  rq_init_comm_if_connected(9, "1")
  rq_init_comm_if_connected(2, "2")
  rq_init_comm_if_connected(3, "3")
  rq_init_comm_if_connected(4, "4")
  rq_print_connected_grippers()
  rq_gripper_communication_thread = run rq_gripper_communication()
  set_closed_norm(97.6470588235294, "1")
  set_open_norm(1.1764705882352942, "1")
  set_closed_mm(0.0, "1")
  set_open_mm(53.0, "1")
  set_closed_norm(100.0, "2")
  set_open_norm(0.0, "2")
  set_closed_mm(0.0, "2")
  set_open_mm(50.0, "2")
  set_closed_norm(100.0, "3")
  set_open_norm(0.0, "3")
  set_closed_mm(0.0, "3")
  set_open_mm(50.0, "3")
  set_closed_norm(100.0, "4")
  set_open_norm(0.0, "4")
  set_closed_mm(0.0, "4")
  set_open_mm(50.0, "4")
  rq_current_limit_enabled = False
  while(not rq_gripper_communication_thread_started):
      sleep(0.008)
  end
  # end: URCap Installation Node
  step_count_126a9c52_0873_4ea5_a9d9_3503bc14fb30 = 0.0
  thread Step_Counter_Thread_0450802b_b3f4_44ca_aa13_af17d282832f():
    while (True):
      step_count_126a9c52_0873_4ea5_a9d9_3503bc14fb30 = step_count_126a9c52_0873_4ea5_a9d9_3503bc14fb30 + 1.0
      sync()
    end
  end
  run Step_Counter_Thread_0450802b_b3f4_44ca_aa13_af17d282832f()
  global TMR_Barcode=0
  global TMR_Barcode_is_counting=False
  thread Timer_Thread():
    while (True):
      if (TMR_Barcode_is_counting):
        TMR_Barcode = TMR_Barcode + get_steptime()
      end
      sync()
    end
  end
  run Timer_Thread()
  $ 2 "BeforeStart"
  $ 3 "Before start"
  $ 4 "Script: SCRIPT Transitions V6.6.script"
  #*****************************************************
  # customer          :   INTERNAL
  # project name      :
  #****************************************************
  # controller        :   UR
  # software          :   5.13
  #****************************************************
  # author            :   P. Koehnke
  # Copyright (c)     :   United Robotics Group
  #                       An der Riede 2
  #                       28816 Stuhr
  #                       Germany
  #****************************************************
  # description       :   transition between workareas
  # version:      	:   1.2
  # created           :   28.02.2024
  # updated           :
  #****************************************************
  # modifications     :
  #
  # date              :
  # name              :
  # reason            :
  #****************************************************

  ######################### further development #########################
  #   - that the robot can switch the configuration, if necessary
  #   - introduction of structs
  #######################################################################

  ######################### to be adjusted #########################
  local WORKAREA_1 = [-0.280,-0.680,-0.001, 0.280, 0.100, 1.000]    # workarea 1 (platform)
  local WORKAREA_2 = [-1.000,-1.000,-1.000,-0.290, 0.100, 1.000]    # workarea 2 (front right)
  local WORKAREA_3 = [-1.000, 0.100,-1.000, 0.000, 1.000, 1.000]    # workarea 3 (back right)
  local WORKAREA_4 = [ 0.000, 0.100,-1.000, 1.000, 1.000, 1.000]    # workarea 4 (back left)
  local WORKAREA_5 = [ 0.290,-1.000,-1.000, 1.000, 0.100, 1.000]    # workarea 5 (front left)
  local WORKAREA_6 = [-0.290,-1.000,-1.000, 0.290,-0.560, 1.000]    # workarea 6 (front front)
  local WORKAREA_7 = [0,0,0,0,0,0]    # reserved
  local WORKAREA_8 = [0,0,0,0,0,0]    # reserved
  local WORKAREA_9 = [0,0,0,0,0,0]    # reserved
  local WORKAREA_10 = [0,0,0,0,0,0]   # reserved

  local PSE_WA_1 = p[ 0.000,-0.450, 0.300, 0.000, 0.000, 0.000]
  local PSE_WA_2 = p[-0.300,-0.300, 0.300, 0.000, 0.000, d2r(-90)]
  local PSE_WA_3 = p[-0.300, 0.300, 0.300, 0.000, 0.000, d2r(-135)]
  local PSE_WA_4 = p[ 0.300, 0.300, 0.300, 0.000, 0.000, d2r(135)]
  local PSE_WA_5 = p[ 0.300,-0.300, 0.300, 0.000, 0.000, d2r(90)]
  local PSE_WA_6 = p[ 0.000,-0.600, 0.300, 0.000, 0.000, 0.000]       # reserved
  local PSE_WA_7 = p[ 0.000, 0.000, 0.000, 0.000, 0.000, 0.000]       # reserved
  local PSE_WA_8 = p[ 0.000, 0.000, 0.000, 0.000, 0.000, 0.000]       # reserved
  local PSE_WA_9 = p[ 0.000, 0.000, 0.000, 0.000, 0.000, 0.000]       # reserved
  local PSE_WA_10 = p[ 0.000, 0.000, 0.000, 0.000, 0.000, 0.000]      # reserved

  global JNT_HOME = [-1.23163,-1.29627,-1.86552,-1.55102, 1.57761, 1.910]
  local JNT_STANDARD_C1 = [ 1.57,-1.57, 1.57,-1.57,-1.57,0]
  local JNT_STANDARD_C2 = [-1.57,-1.57,-1.57,-1.57, 1.57,0]
  local YAW_MIN_DEG = -110
  local YAW_MAX_DEG = 110
  local DISTANCE_TO_CLEARANCE = 0.300
  local RADIUS_HELPER_POSES = 0.300
  local RADIUS_TRANSITION_POSES = 0.400
  local workareas = [WORKAREA_1, WORKAREA_2, WORKAREA_3, WORKAREA_4, WORKAREA_5, WORKAREA_6, WORKAREA_7, WORKAREA_8, WORKAREA_9, WORKAREA_10]
  local poses = [PSE_WA_1, PSE_WA_2, PSE_WA_3, PSE_WA_4, PSE_WA_5, PSE_WA_6, PSE_WA_7, PSE_WA_8, PSE_WA_9, PSE_WA_10]

  ######################### end of adjustment #########################

  local pi = 3.14159265
  local axis_config_current = 0
  local axis_config_new = 0
  local workarea_current = 0
  local workarea_new = 0
  global reverse_rotation = False

  def create_transition_pose():
      return struct(crt = p[0,0,0,0,0,0], jnt = [0,0,0,0,0,0], q = [0,0,0,0,0,0], yaw_too_base = 0.0)
  end

  local pose_start = create_transition_pose()
  local pose_help = create_transition_pose()
  local pose_target = create_transition_pose()
  local pose = create_transition_pose()

  def init_home_by_cartesian_pose(pose):
      # check given pose for reachability for the corresponding axis config
      global pose_inv_tcp = pose_inv(get_tcp_offset())
      global pose_tcp_offset = get_tcp_offset()
      global pose_home = pose_trans(pose, pose_inv_tcp)

      if check_current_axis_config() == 1:
          if get_inverse_kin_has_solution(pose_home, qnear=JNT_STANDARD_C1, tcp=p[0,0,0,0,0,0]):
              JNT_HOME = get_inverse_kin(pose_home, qnear=JNT_STANDARD_C1, tcp=p[0,0,0,0,0,0])
          end
      elif check_current_axis_config() == 2:
          if get_inverse_kin_has_solution(pose_home, qnear=JNT_STANDARD_C2, tcp=p[0,0,0,0,0,0]):
              JNT_HOME = get_inverse_kin(pose_home, qnear=JNT_STANDARD_C2, tcp=p[0,0,0,0,0,0])
          end
      end
  end

  def get_tool_free_pose(pose_ref=get_actual_tcp_pose(), dir=[0,0,0], move_in_base_frame=False):
      # get a recovery pose
      # dir is providing the direction and distance in X, Y and Z
      # if 'move_in_base_frame' is set, dir will be interpreted as absolute values for a movement in base frame

      local pose_target = pose_ref
      local i = 0

      if (move_in_base_frame):
          while (i<3):
              # move only,
              # if the demanded position is bigger than zero and the current position is below the demanded one or
              # if the demanded position is smaller than zero and the current position is above the demanded one
              if ((dir[i]>0 and pose_ref[i]<dir[i]) or (dir[i]<0 and pose_ref[i]>dir[i])):
                  pose_target[i] = dir[i]
              end
              i = i + 1
          end
      else:
          pose_target = pose_trans(pose_ref, p[dir[0], dir[1], dir[2], 0, 0, 0])
      end

      return pose_target
  end

  def check_workarea(reference_pose):
      # the actual TCP position is compared to predefined areas (cubic) to determine in which area the robot arm is
      # a workarea is defined as a list of coordinates, where the first 3 values are X, Y, and Z with the smallest values and
      # the next 3 values specify X, Y and Z for the biggest values

      local data_size = size(workareas)
      local i = 0
      local size_workarea = p[0,0,0,0,0,0]
      local pose_workarea = p[0,0,0,0,0,0]

      while (i < data_size[0]):
          pose_workarea = pose_trans(inv(p[workareas[i, 0], workareas[i, 1], workareas[i, 2], 0, 0, 0]), reference_pose)
          size_workarea = pose_sub(p[workareas[i, 3], workareas[i, 4], workareas[i, 5], 0, 0, 0], p[workareas[i, 0], workareas[i, 1], workareas[i, 2], 0, 0, 0])
          if  ((pose_workarea[0]>0 and pose_workarea[0]<size_workarea[0]) and
              (pose_workarea[1]>0 and pose_workarea[1]<size_workarea[1]) and
              (pose_workarea[2]>0 and pose_workarea[2]<size_workarea[2])):
              return i + 1
          end
          i = i + 1
      end
      return 0
  end

  def check_current_axis_config():
      # function determnines, if the arm is oriented in one or the other configuration.
      # it means, that the ellbow joint is flipped and so are the wrist joints.

      local jnt_current = get_actual_joint_positions()

      # ellbow has positiv angle
      if (jnt_current[2]> 0):
          return 1
      # ellbow has negativ angle
      elif (jnt_current[2]< 0):
          return 2
      # angle is 0
      else:
          return 0
      end
  end

  def switch_axis_config(axis_config):
      # function to switch betwwen the axis configuration 1 and 2.

      if (axis_config == 1):
          return 2
      elif (axis_config ==2):
          return 1
      end
  end

  def get_transition_pose_by_workarea(workarea, axis_config):
      # get the correspondig pose from the list of poses

      pose.crt = poses[workarea-1]
      pose.yaw_too_base = get_yaw_too_base(pose.crt)
      pose.q = get_actual_joint_positions()

      if get_inverse_kin_has_solution(pose.crt, qnear=pose.q):
          pose.jnt = get_inverse_kin(pose.crt, qnear=pose.q)
      else:
          popup("no solution found for the transition pose", blocking= True)
      end

      return pose
  end

  def get_transition_pose_by_reference_pose(ref, radius, axis_config):
      # get the correspondig pose from the list of poses

      pose.yaw_too_base = get_yaw_too_base(ref)
      pose.q = get_actual_joint_positions()

      # get coordinates of the circle with the same angle as the given pose to the
      if ref == p[0,0,0,0,0,0]:
          pose.q = JNT_HOME
          pose.jnt = JNT_HOME
          pose.crt = get_forward_kin(pose.jnt)
          return pose
      else:
          pose.crt = p[
              radius * cos(pose.yaw_too_base-pi/2),
              radius * sin(pose.yaw_too_base-pi/2),
              DISTANCE_TO_CLEARANCE,
              0,
              0,
              pose.yaw_too_base + get_locked_yaw()]
      end

      if get_inverse_kin_has_solution(pose.crt, qnear=pose.q):
          pose.jnt = get_inverse_kin(pose.crt, qnear=pose.q)
      else:
          popup("no solution found for the transition pose", blocking= True)
      end

      return pose
  end

  def get_transition_pose_by_yaw(yaw, radius, axis_config):

      pose.yaw_too_base = yaw
      pose.q = get_actual_joint_positions()
      pose.crt = p[
          radius * cos(yaw-pi/2),
          radius * sin(yaw-pi/2),
          DISTANCE_TO_CLEARANCE,
          0,
          0,
          yaw + get_locked_yaw()]

      if get_inverse_kin_has_solution(pose.crt, qnear=pose.q):
          pose.jnt = get_inverse_kin(pose.crt, qnear=pose.q)
      else:
          popup("no solution found for the transition pose", blocking= True)
      end

      return pose
  end

  def get_rounded_mm(value):
      if (value < 0):
          return ceil(value*1000)
      elif (value >= 0):
          return floor(value*1000)
      end
  end

  def get_yaw_too_base(pose):
      # get the yaw relative to the base frame
      local pose_x_mm = 0
      local pose_y_mm = 0
      local yaw = 0

      pose_x_mm = get_rounded_mm(pose[0])
      pose_y_mm = get_rounded_mm(pose[1])

      if (pose_x_mm == 0 and pose_y_mm < 0):
          yaw = 0
      elif (pose_x_mm == 0 and pose_y_mm > 0):
          yaw = pi
      elif (pose_x_mm < 0 and pose_y_mm == 0):
          yaw = -pi/2
      elif (pose_x_mm > 0 and pose_y_mm == 0):
          yaw = pi/2
      else:
          yaw = atan2(pose[0], pose[1])
          if (-pi < yaw) and (yaw < 0):
              yaw = - yaw - pi
          elif (0 < yaw) and (yaw < pi):
              yaw = - yaw + pi
          end
      end
      return yaw
  end

  def adjust_axis_rotation(pose):

      if (0 > pose.yaw_too_base) and (pose.yaw_too_base > d2r(YAW_MIN_DEG)):
          if (pose.jnt[0] > JNT_HOME[0]):
              # calculated axis angle is in the wrong value range
              if axis_config_current == 1:
                  pose.q[0] = JNT_STANDARD_C1[0]
              elif axis_config_current == 2:
                  pose.q[0] = JNT_STANDARD_C2[0]
              end
              reverse_rotation = True
          end
      elif (0 < pose.yaw_too_base) and (pose.yaw_too_base < d2r(YAW_MAX_DEG)):
          if (pose.jnt[0] < JNT_HOME[0]):
              if axis_config_current == 1:
                  pose.q[0] = JNT_STANDARD_C1[0]
              elif axis_config_current == 2:
                  pose.q[0] = JNT_STANDARD_C2[0]
              end
              reverse_rotation = True
          end
      elif (pose.jnt[0] < -2 * pi):
          if axis_config_current == 1:
              pose.q[0] = JNT_STANDARD_C1[0]
          elif axis_config_current == 2:
              pose.q[0] = JNT_STANDARD_C2[0]
          end
          reverse_rotation = True
      elif (pose.jnt[0] > 2 * pi):
          if axis_config_current == 1:
              pose.q[0] = JNT_STANDARD_C1[0]
          elif axis_config_current == 2:
              pose.q[0] = JNT_STANDARD_C2[0]
          end
          reverse_rotation = True
      end
      return pose.q[0]
  end

  def adjust_transition_poses(pose_identifier, keep_rxry=False):
      # adjust the orientation of the transition poses by determining the the current orientation

      local pose_current = get_actual_tcp_pose()
      local jnt_current = get_actual_joint_positions()
      local rpy_current = rotvec2rpy([pose_current[3],pose_current[4],pose_current[5]])
      local rotvec_new = [0,0,0]

      if (pose_identifier == "start"):
          pose = pose_start
      elif (pose_identifier == "target"):
          pose = pose_target
          pose.q[0] = adjust_axis_rotation(pose)
      elif (pose_identifier == "helper"):
          pose = pose_help
      end

      if keep_rxry:
          rotvec_new = rpy2rotvec([rpy_current[0], rpy_current[1], pose.yaw_too_base + get_locked_yaw()])
          pose.crt = p[pose.crt[0], pose.crt[1], pose.crt[2], rotvec_new[0], rotvec_new[1], rotvec_new[2]]

          # adjust preferred joint angles ot the current ones
          pose.q[3] = jnt_current[3]
          pose.q[4] = jnt_current[4]
          pose.q[5] = jnt_current[5]
      end

      if get_inverse_kin_has_solution(pose.crt, qnear=pose.q) and is_within_safety_limits(pose.crt):
          pose.jnt = get_inverse_kin(pose.crt, qnear=pose.q)
      else:
          popup(str_cat("no solution for ", pose_identifier), error=True, blocking=True)
      end
      return pose.jnt
  end

  def get_locked_yaw():
      local pose_current = get_actual_tcp_pose()
      local rpy_current = rotvec2rpy([pose_current[3],pose_current[4],pose_current[5]])
      local rotvec_new = rpy2rotvec([rpy_current[0], rpy_current[1], get_yaw_too_base(pose_current)])
      local pose_reference = p[pose_current[0], pose_current[1], pose_current[2], rotvec_new[0], rotvec_new[1], rotvec_new[2]]
      local pose_to_reference = pose_trans(pose_inv(pose_reference), pose_current)

      return pose_to_reference[5]
  end

  def get_helper_yaw():
      local yaw = 0

      yaw = (pose_start.yaw_too_base + pose_target.yaw_too_base) / 2

      if reverse_rotation and
          ((pose_start.yaw_too_base < 0 and
          pose_target.yaw_too_base < 0) or
          (pose_start.yaw_too_base > 0 and
          pose_target.yaw_too_base > 0)):
            yaw = flip_yaw(yaw)
      elif (pose_start.yaw_too_base < 0 and
            pose_start.yaw_too_base < d2r(YAW_MIN_DEG)) and
            (pose_target.yaw_too_base > 0 and
            pose_target.yaw_too_base > d2r(YAW_MAX_DEG)):
              yaw = flip_yaw(yaw)
      elif (pose_start.yaw_too_base > 0 and
            pose_start.yaw_too_base > d2r(YAW_MAX_DEG)) and
            (pose_target.yaw_too_base < 0 and
            pose_target.yaw_too_base < d2r(YAW_MIN_DEG)):
              yaw = flip_yaw(yaw)
      end
      return yaw
  end

  def flip_yaw(yaw):
      # flips the given yaw 180 degree around
      if (yaw < 0):
          return yaw + pi
      elif (yaw > 0):
          return yaw - pi
      end
  end

  def clear_poses():
      pose = create_transition_pose()
      pose_start = create_transition_pose()
      pose_help = create_transition_pose()
      pose_target = create_transition_pose()
  end

  def do_transition(reference_pose=p[0,0,0,0,0,0], mode=2, keep_rxry=False, a=1.4, v=1.05, r=0.100):
      # the robot will evaluate the current and target workarea
      # after that, the robot will move between the workareas automatically.
      # parameters:
      # reference_pose:   a pose/frame were the robot should work next. If nothing is given, base frame will be used as target
      # keep_rxry:        if true, the robot will keep the orientation of the tool during the movement

      ################# checking #################
      axis_config_current = check_current_axis_config()           # 0: unknown, 1: config 1, 2: config 2
      workarea_current = check_workarea(get_actual_tcp_pose())    # between 0 and the amount of defined workareas
      workarea_new = check_workarea(reference_pose)               # between 0 and the amount of defined workareas
      reverse_rotation = False

      if (workarea_current != 0 and workarea_new != 0) and (workarea_current != workarea_new) or (reference_pose == p[0,0,0,0,0,0]):
          ################# get axisvalues #################
          if (mode == 1):
              pose_start = get_transition_pose_by_workarea(workarea_current, axis_config_current)
              pose_target = get_transition_pose_by_workarea(workarea_new, axis_config_current)
          elif (mode == 2):
              pose_start = get_transition_pose_by_reference_pose(get_actual_tcp_pose(), RADIUS_TRANSITION_POSES, axis_config_current)
              pose_target = get_transition_pose_by_reference_pose(reference_pose, RADIUS_TRANSITION_POSES, axis_config_current)
          end

          ################# adjustments #################
          pose_start.jnt = adjust_transition_poses("start", keep_rxry)
          pose_target.jnt = adjust_transition_poses("target", keep_rxry)

          if (pose_start.crt[1] < 0 and pose_target.crt[1] > 0) or (pose_start.crt[1] > 0 and pose_target.crt[1] < 0):
              pose_help = get_transition_pose_by_yaw(get_helper_yaw(), RADIUS_HELPER_POSES, axis_config_current)
              pose_help.jnt = adjust_transition_poses("helper", keep_rxry)
          end

          ################# movements #################
          if (pose_help.jnt != [0,0,0,0,0,0]):
              if point_dist(get_actual_tcp_pose(), pose_start.crt) > r and point_dist(pose_start.crt, pose_help.crt) > r:
                  movej(pose_start.jnt, a=a, v=v, r=r)
                  if (point_dist(pose_start.crt, pose_help.crt) > r) and (point_dist(pose_target.crt, pose_help.crt) > r):
                      movej(pose_help.jnt, a=a, v=v, r=r)
                  end
              end
          else:
              if point_dist(get_actual_tcp_pose(), pose_start.crt) > r and point_dist(pose_start.crt, pose_target.crt) > r:
                  movej(pose_start.jnt, a=a, v=v, r=r)
              end
          end
          movej(pose_target.jnt, a=a, v=v)
      else:
          # define error
      end

      ################# checking #################
      axis_config_current = check_current_axis_config()           # 0: unknown, 1: config 1, 2: config 2
      workarea_current = check_workarea(get_actual_tcp_pose())    # between 0 and the amount of defined workareas
      clear_poses()
  end
  $ 5 "Script: SCRIPT Utility V5.4.script"
  #*****************************************************
  # customer          :   tbd
  # project name      :   tbd
  #****************************************************
  # controller        :
  # software          :
  #****************************************************
  # author            :   P. Koehnke (+49 1628859904; p.koehnke@unitedrobotics.group)
  # Copyright (c)     :   United Robotics Group Health and Food GmbH
  #                       An der Riede 2
  #                       28816 Stuhr
  #                       Germany
  #****************************************************
  # description       :   utility programs for the application
  # version:      	:   3.1
  # created           :   30.01.2023
  # updated           :
  #****************************************************
  # modifications     :   get_tool_free_pose_2(), get_index_from_list()
  #
  # date              :   05.01.2024
  # name              :   PK
  # reason            :
  #****************************************************

  def found_in_matrix(data, req_id, req_idx):
      local id = -1
      local dimensions = size(data)
      local loop_dataset = 0

      while (id != req_id and loop_dataset < dimensions[0]):
          id = data[loop_dataset, 0]
          if (id == req_id):
              return data[loop_dataset, req_idx]
          else:
              loop_dataset = loop_dataset + 1
          end
      end
  end

  def found_in_list(value, list):
      local idx = 0

      while (idx < length(list)):
          if (value == list[idx]):
              return True
          end
          idx = idx + 1
      end
      return False
  end

  def get_index_from_list(list, value = -1):
      local idx = 0

      while (idx < length(list)):
          if (value == -1):
              if (list[idx] != 0):
                  return idx
              end
          else:
              if (list[idx] == value):
                  return idx
              end
          end
          idx = idx + 1
      end
      return -1
  end

  def find_object_by_type(list, type=0):
      local object = list[0]
      local i = 0

      while i < length(list):
          object = list[i]
          if object.type == type:
              return object
          end
          i = i + 1
      end
  end

  def pose_RPY2RotVec(pose):
      local rotvec = rpy2rotvec([d2r(pose[3]), d2r(pose[4]), d2r(pose[5])])
      return p[pose[0], pose[1], pose[2], rotvec[0], rotvec[1], rotvec[2]]
  end

  def pose_RotVec2RPY(pose):
      local rpy = rotvec2rpy([pose[3], pose[4], pose[5]])
      return p[pose[0], pose[1], pose[2], r2d(rpy[0]), r2d(rpy[1]), r2d(rpy[2])]
  end

  def swivel(frame_ref, angles = [0, 0, 0], pose = p[0, 0, 0, 0, 0, 0]):

      local rpy_ref = [0, 0, 0]
      local rpy_new = [0, 0, 0]
      local rotvec_new = [0, 0, 0]
      local pose_from = p[0, 0, 0, 0, 0, 0]
      local pose_to = p[0, 0, 0, 0, 0, 0]
      local i = 0

      if (pose == p[0, 0, 0, 0, 0, 0]):
          pose_to = pose_trans(pose_inv(frame_ref), get_actual_tcp_pose())
      else:
          pose_to = pose
      end

      rpy_ref = rotvec2rpy(frame_ref[3], frame_ref[4], frame_ref[5])

      while (i < 3):
          rpy_new[i] = rpy_ref[i] + d2r(angles[i])
          i = i + 1
      end

      rotvec_new = rpy2rotvec(rpy_new)
      pose_from = p[0, 0, 0, rotvec_new[0], rotvec_new[1], rotvec_new[2]]
      pose_to = p[pose_to[0], pose_to[1], pose_to[2], rotvec_new[0], rotvec_new[1], rotvec_new[2]]

      return pose_trans(pose_from, pose_to)
  end

  def get_random_pose(pose_ref, mode = "", range_max = [0, 0, 0]):
      # modi: "cubic", "rotation"
      # getting a random pose in the x/y-plane. range can be set for each
      # translation and rotation.
      local rpy_random = [0, 0, 0]
      local rotvec_random = [0, 0, 0]
      local pose_random = pose_ref
      local i = 0

      if (mode == "cubic"):
          # cubic mode: random pose takes only x, y and z
          i = 0
          while (i < 3):
              pose_random[i] = pose_ref[i] + range_max[i] * (random() - 0.5)
              i = i + 1
          end
          return pose_random

      elif (mode == "rotation"):
          i = 0
          while (i < 3):
              rpy_random[i] = d2r(range_max[i]) * (random() - 0.5)
              i = i + 1
          end
          rotvec_random = rpy2rotvec(rpy_random)
          pose_random = pose_trans(p[0, 0, 0, rotvec_random[0], rotvec_random[1], rotvec_random[2]], pose_ref)
          return pose_random

      else:
          # unknown mode, return pose_ref
          return pose_ref
      end
  end

  def get_pattern_pos_rectangle(counter, direction, pattern, patterninc = [0, 0], patternsize = [0, 0]):
      # defines the position inside a rectangular pattern
      # pattern describes, how many objects are in x-direction and how many in y-direction [x, y]
      # patternsize will give the total length of each direction [x, y]
      local X_Fac = 0
      local Y_Fac = 0
      local max = pattern[0] * pattern[1]
      local i = 0

      if (1 > counter or counter > max):
          counter = 1
      end

      if pattern[0] == 0:
          pattern[0] = 1
      end

      if pattern[1] == 0:
          pattern[1] = 1
      end

      if (direction == "Y" or direction == "y"):
          X_Fac = floor((counter - 1) / pattern[1])
          Y_Fac = (counter - 1) % pattern[1]
      elif (direction == "X" or direction == "x"):
          X_Fac = (counter - 1) % pattern[0]
          Y_Fac = floor((counter - 1) / pattern[0])
      end

      if patternsize != [0, 0]:
          while i < 2:
              if pattern[i] > 1:
                  patterninc[i] = patternsize[i] / (pattern[i] - 1)
              end
              i = i + 1
          end
      end

      return p[X_Fac * patterninc[0], Y_Fac * patterninc[1], 0, 0, 0, 0]
  end

  def get_pattern_pos_circle(counter, radius, angle, direction, pattern, patternsize = [0, 0]):
      # get the patternpos for a circular pattern through a counter
      # need the radius and the angle in radiants
      local X_Fac = 0
      local Y_Fac = 0
      local rad_bow = 0
      local radius_cal = 0
      local ref = p[0, 0, 0, 0, 0, 0]

      if pattern[0] == 0:
          pattern[0] = 1
      end

      if pattern[1] == 0:
          pattern[1] = 1
      end

      if (direction == "Y" or direction == "y"):
          X_Fac = floor((counter - 1) / pattern[1])
          Y_Fac = (counter - 1) % pattern[1]
      elif (direction == "X" or direction == "x"):
          X_Fac = (counter - 1) % pattern[0]
          Y_Fac = floor((counter - 1) / pattern[0])
      end

      # the opening angle will be calculated in x-direction
      # works only between -90 and 90 degree
      if pattern[0] > 1:
          rad_bow = - angle / (pattern[0] - 1) * X_Fac + angle / 2
      end

      if (counter % 2 == 0 and pattern[1] > 1):
          radius_cal = radius - patternsize[1] / (pattern[1])
      else:
          radius_cal = radius + patternsize[1] / (pattern[1])
      end
      ref = p[0, radius_cal, 0, 0, 0, 0]

      return p[ref[0] * cos(rad_bow) - ref[1] * sin(rad_bow), (ref[0] * sin(rad_bow) + ref[1] * cos(rad_bow)) - radius, 0, 0, 0, 0]
  end

  def get_pattern_counter(pose, direction, pattern, patterninc = [0, 0], patternsize = [0, 0]):
      # returns the counter for a pattern from a given cartesian pose
      local patternpose = p[pose[0], pose[1], 0, 0, 0, 0]
      local X_Fac = 0
      local Y_Fac = 0
      local i = 0

      if patternsize != [0, 0]:
          while i < 2:
              if pattern[i] > 1:
                  patterninc[i] = patternsize[i] / (pattern[i] - 1)
              else:
                  pattern[i] = 0
              end
              i = i + 1
          end
      end

      # calculation of the counter in the desired axis-direction
      if (direction == "x" or direction == "X"):
          if patterninc[0] > 0:
              X_Fac = ceil((patternpose[0] + patterninc[0] / 2) / patterninc[0])
              if X_Fac < 0:
                  X_Fac = 0
              end
          end
          if patterninc[1] > 0:
              Y_Fac = floor((patternpose[1] + patterninc[1] / 2) / patterninc[1])
              if Y_Fac < 0:
                  Y_Fac = 0
            end
          end
          return Y_Fac * pattern[0] + X_Fac
      elif (direction == "y" or direction == "Y"):
          if patterninc[0] > 0:
              X_Fac = floor((patternpose[0] + patterninc[0] / 2) / patterninc[0])
          end
          if patterninc[1] > 0:
              Y_Fac = ceil((patternpose[1] + patterninc[1] / 2) / patterninc[1])
          end
          return X_Fac * pattern[1] + Y_Fac
      end
  end

  def get_plc_reg(mod_sig_name):
      return integer_to_binary_list(modbus_get_signal_status(mod_sig_name))
  end

  def set_plc_reg(mod_sig_name, mod_sig_list):
      modbus_set_output_register(mod_sig_name, binary_list_to_integer(mod_sig_list), False)
  end

  def check_decapping(offset = 0, timeout = 5, abort = False):
      # checken, ob der Deckel schon ab ist
      local start = get_actual_tcp_pose()
      local current_offset = 0
      local timecounter = 0
      while (current_offset < offset and not abort):
          current_offset = pose_dist(start, get_actual_tcp_pose())
          timecounter = timecounter + 1
          if (timecounter * 0.5 == timeout):
              break
          end
          sleep(0.5)
      end
      stopl(0.5)
  end

  def check_capping(torque = 0):
      # checken, wann der Deckel verschraubt ist
      force_mode(get_actual_tcp_pose(), [0, 0, 1, 0, 0, 0], [0, 0, -2.0, 0, 0, 0], 2, [0, 0, 0.100, 0, 0, 0])
  end

  def is_reachable(frame, poses, offsets = [0, 0, 0]):
      local idx = 0
      local pose = p[0, 0, 0, 0, 0, 0]

      while (idx < length(poses)):
          pose = poses[idx]
          pose[0] = pose[0] + offsets[0]
          pose[1] = pose[1] + offsets[1]
          pose[2] = pose[2] + offsets[2]

          if pose != p[0, 0, 0, 0, 0, 0]:
              if (not get_inverse_kin_has_solution(pose_trans(frame, pose))):
                  textmsg(str_cat(str_cat("Pose ", to_str(idx + 1)), " is not reachable"))
                  return False
              end
          end
          idx = idx + 1
      end
      return True
  end

  def is_within_limits(frame, poses, offsets = [0, 0, 0]):
      local idx = 0
      local pose = p[0, 0, 0, 0, 0, 0]

      while (idx < length(poses)):
          pose = poses[idx]
          pose[0] = pose[0] + offsets[0]
          pose[1] = pose[1] + offsets[1]
          pose[2] = pose[2] + offsets[2]

          if is_reachable(frame = frame, poses = poses, offsets = offsets):
              if (not is_within_safety_limits(get_inverse_kin(pose_trans(frame, pose), get_actual_joint_positions()))):
                  textmsg(str_cat(str_cat("Pose ", to_str(idx + 1)), "is out of joint limits"))
                  return False
              else:
                  idx = idx + 1
              end
          else:
              return False
          end
      end
      return True
  end
  $ 6 "Script: SCRIPT Objects V0.1.script"
  #*****************************************************
  # customer          :   INTERNAL
  # project name      :
  #****************************************************
  # controller        :   UR
  # software          :   5.17.3
  #****************************************************
  # author            :   P. Koehnke
  # Copyright (c)     :   United Robotics Group
  #                       An der Riede 2
  #                       28816 Stuhr
  #                       Germany
  #****************************************************
  # description       :   object database
  # version:      	:   0.1
  # created           :   09.10.2024
  # updated           :
  #****************************************************
  # modifications     :
  #
  # date              :
  # name              :
  # reason            :
  #****************************************************

  def create_object_2(id=0, name="", type=0, dimension=struct(length=0, width=0, height=0, diameter=0), gripper_offset=p[0,0,0,0,0,0]):
      return struct(id=id, name=name, type=type, dimension=dimension, gripper_offset=gripper_offset)
  end

  OBJ = create_object_2()
  OBJs = make_list(0, create_object_2(), 50)

  OBJs.append(create_object_2(id=1, name="rack centrifuge", type=1, dimension=struct(length=0, width=0, height=0.106, diameter=0.020), gripper_offset=p[0,0,0.095,0,0,2.356]))
  OBJs.append(create_object_2(id=2, name="sample tube 1", type=2, dimension=struct(length=0, width=0, height=0.106, diameter=0.015), gripper_offset=p[0,0,0.060,0,0,0]))

  def create_jig_2(id=0, name="", type=0, capacity=0, jig_offset=p[0,0,0,0,0,0]):
      # iformation about used jigs
      return struct(id=id, name=name, type=type, capacity=capacity, jig_offset=jig_offset)
  end

  JIG2 = create_jig_2()
  JIGs = make_list(0, create_jig_2(), 10)

  JIGs.append(create_jig_2(id=1, name="3FG", type=1, capacity=1, jig_offset=p[0,0,0,0,0,0]))
  JIGs.append(create_jig_2(id=2, name="jig input", type=2, capacity=1, jig_offset=p[0,0,0,0,0,-3.927]))
  JIGs.append(create_jig_2(id=3, name="jig output", type=3, capacity=1, jig_offset=p[0,0,0,0,0,0.78]))
  JIGs.append(create_jig_2(id=4, name="jig centrifuge racks", type=4, capacity=4, jig_offset=p[0,0,0,0,0,-3.9162]))
  $ 7 "Script: 001 SCRIPT Errors and Warnings Deifnes V0.2.script"

  #*****************************************************
  # customer          :   UK Essen
  # project name      :   P1132
  #****************************************************
  # controller        :
  # software          :
  #****************************************************
  # author            :   E.Petrichenko
  # Copyright (c)     :   United Robotics Group Health and Food GmbH
  #                       An der Riede 2
  #                       28816 Stuhr
  #                       Germany
  #****************************************************
  # description       :   centrifuge actions for the application
  # version:      	:   0.1
  # created           :   22.08.2024
  # updated           :
  #****************************************************
  # modifications     :
  #
  # date              :
  # name              :
  # reason            :
  #****************************************************


  #################################### VARIABLES DEFINITIONS ###################################

  ERROR_POSE_NOT_REACHABLE = 1002
  ERROR_ROBOT_ARM_NOT_IN_HOME_POSE = 1006
  ERROR_NO_OBJECT_TO_PICK = 1010
  ERROR_NOT_DOCKED = 2003
  ERROR_NOT_REACHABLE_TARGET = 2007
  ERROR_CHARGING_NOT_STARTED = 2008
  ERROR_AMR_WRONG_MODE = 2009
  ERROR_UNKNOWN_POSE = 2010
  ERROR_NO_LANDMARK = 3002
  ERROR_WRONG_ORDER = 4002
  ERROR_CENTRIFUGE_CONNECTION = 5001
  ERROR_CENTRIFUGE_POWER = 5002
  ERROR_CENTRIFUGE = 5003
  ERROR_CENTRIFUGE_LID = 5004
  ERROR_CANNOT_OPEN_HATCH = 5006
  ERROR_CANNOT_CLOSE_HATCH = 5008
  ERROR_CANNOT_ROTATE = 5010
  ERROR_CANNOT_START = 5011
  ERROR_WRONG_KEY_POSE = 5012
  ERROR_MISSIING_CENTRACK = 5013

  WARNING_POSE_NOT_REACHABLE = 1002
  WARNING_BATTERY_LEVEL = 2002
  WARNING_NOT_REACHABLE_TARGET = 2007


  ERROR = struct(
      FLAG = False,
      ID = 0,
      MSG = "")

  WARNING = struct(
      FLAG = False,
      ID = 0,
      MSG = "")


  #################################### FUNCTIONS ###################################

  def set_error(error_id):
      ERROR.ID = error_id
      if (ERROR.ID == 0):
          ERROR.FLAG = False
          ERROR.MSG = ""
      else:
          ERROR.FLAG = True
          if(ERROR.ID == ERROR_POSE_NOT_REACHABLE):
              ERROR.MSG = "Pose is not reachable"
          elif(ERROR.ID == ERROR_NO_OBJECT_TO_PICK):
              ERROR.MSG = "No object to pick"
          elif(ERROR.ID == ERROR_NO_LANDMARK):
              ERROR.MSG = "No landmark detected"
          elif(ERROR.ID == ERROR_ROBOT_ARM_NOT_IN_HOME_POSE):
              ERROR.MSG = "Robot arm cannot go to home pose"
          elif(ERROR.ID == ERROR_AMR_WRONG_MODE):
              ERROR.MSG = "AMR is in the wrong mode"
          elif(ERROR.ID == ERROR_NOT_DOCKED):
              ERROR.MSG = "Could not dock to the charger"
          elif(ERROR.ID == ERROR_NOT_REACHABLE_TARGET):
              ERROR.MSG = "Could not reach the target"
          elif(ERROR.ID == ERROR_CHARGING_NOT_STARTED):
              ERROR.MSG = "Could not start charging"
          elif(ERROR.ID == ERROR_UNKNOWN_POSE):
              ERROR.MSG = "Unknown navigation target"
          elif(ERROR.ID == ERROR_CANNOT_OPEN_HATCH):
              ERROR.MSG = "Centrifuge Cannot open the hatch"
          elif(ERROR.ID == ERROR_CENTRIFUGE_CONNECTION):
              ERROR.MSG = "Cannot reach centrifuge"
          elif (ERROR.ID == ERROR_CANNOT_CLOSE_HATCH):
              ERROR.MSG = "Centrifuge Cannot close the hatch"
          elif (ERROR.ID == ERROR_CANNOT_START):
              ERROR.MSG = "Centrifuge Cannot start"
          elif (ERROR.ID == ERROR_CANNOT_ROTATE):
              ERROR.MSG = "Centrifuge Cannot rotate the rotor"
          elif (ERROR.ID == ERROR_WRONG_ORDER):
              ERROR.MSG = "Wrong parameter was recieved"
          elif (ERROR.ID == ERROR_CENTRIFUGE):
              ERROR.MSG = "Centrifuge is in Error"
          elif (ERROR.ID == ERROR_WRONG_KEY_POSE):
              ERROR.MSG = "Key is in the wrong position"
          elif(ERROR.ID == ERROR_MISSIING_CENTRACK):
              ERROR.MSG = "Missing rack for centrifuge set"
          elif(ERROR.ID == ERROR_CENTRIFUGE_POWER):
              ERROR.MSG = "Centrifuge is turned off"
          elif(ERROR.ID == ERROR_CENTRIFUGE_LID):
              ERROR.MSG = "Lid of the centrifuge is opened"
          else:
              ERROR.MSG = "Unknown code"
          end
          textmsg("ERROR:",ERROR)
      end
  end

  def set_warning(warning_id):
      WARNING.ID = warning_id
      if (WARNING.ID == 0):
          WARNING.FLAG = False
          WARNING.MSG = ""
      else:
          WARNING.FLAG = True
          if(WARNING.ID == WARNING_POSE_NOT_REACHABLE):
              WARNING.MSG = "Pose is not reachable"
          elif(WARNING.ID == WARNING_BATTERY_LEVEL):
              WARNING.MSG = "Batery level dropped to a certain level"
          elif(WARNING.ID == WARNING_NOT_REACHABLE_TARGET):
              WARNING.MSG = "Not reachable location of AMR"
          else:
              WARNING.MSG = "Unknown code"
          end
          textmsg("WARNING:",WARNING)
      end
  end


  def reset_error():
    ERROR.ID = 0
    ERROR.FLAG = False
    ERROR.MSG = ""
  end


  def reset_warning():
      WARNING.ID = 0
      WARNING.FLAG = False
      WARNING.MSG = ""
    end
  $ 8 "ITM_ID≔1"
  global ITM_ID=1
  $ 9 "JIG≔2"
  global JIG=2
  $ 10 "JIG_Slot≔3"
  global JIG_Slot=3
  $ 11 "OBJ_Type≔2"
  global OBJ_Type=2
  $ 12 "OBJ_Nbr≔4"
  global OBJ_Nbr=4
  $ 13 "Action≔2"
  global Action=2
  $ 14 "Robot Program"
  $ 15 "PreSettings"
  $ 16 "init poses"
  $ 17 "PSE_A≔p[0,0,0,0,0,0]"
  global PSE_A=p[0,0,0,0,0,0]
  $ 18 "PSE_A_H≔p[0,0,0,0,0,0]"
  global PSE_A_H=p[0,0,0,0,0,0]
  $ 19 "PSE_T≔p[0,0,0,0,0,0]"
  global PSE_T=p[0,0,0,0,0,0]
  $ 20 "PSE_T_H≔p[0,0,0,0,0,0]"
  global PSE_T_H=p[0,0,0,0,0,0]
  $ 21 "PSE_G≔p[0,0,0,0,0,0]"
  global PSE_G=p[0,0,0,0,0,0]
  $ 22 "PSE_G_H≔p[0,0,0,0,0,0]"
  global PSE_G_H=p[0,0,0,0,0,0]
  $ 23 "PSE_R≔p[0,0,0,0,0,0]"
  global PSE_R=p[0,0,0,0,0,0]
  $ 24 "PSE_R_H≔p[0,0,0,0,0,0]"
  global PSE_R_H=p[0,0,0,0,0,0]
  $ 25 "JNT_Q≔[0,0,0,0,0,0]"
  global JNT_Q=[0,0,0,0,0,0]
  $ 26 "JNT_S≔[0,0,0,0,0,0]"
  global JNT_S=[0,0,0,0,0,0]
  $ 27 "Gripping parameters"
  $ 28 "OBJ = find_object_by_type(OBJs, OBJ_Type)"
  OBJ = find_object_by_type(OBJs, OBJ_Type)
  $ 29 "GRP_Open_Pos≔OBJ.dimension.diameter * 1000 + 6"
  global GRP_Open_Pos=OBJ.dimension.diameter * 1000 + 6
  $ 30 "GRP_Offset≔OBJ.gripper_offset"
  global GRP_Offset=OBJ.gripper_offset
  $ 31 "rq_set_force_norm(50)"
   rq_set_force_norm (50)
  $ 32 "rq_set_speed_norm(50)"
   rq_set_speed_norm (50)
  $ 33 "Switch ITM_ID"
  switch_1 = ITM_ID
  $ 34 "Case 1"
  if (1 == switch_1):
    $ 35 "uML"
    $ 36 "JIG2 = find_object_by_type(JIGs, JIG)"
    JIG2 = find_object_by_type(JIGs, JIG)
    $ 37 "JIG_Offset≔JIG2.jig_offset"
    global JIG_Offset=JIG2.jig_offset
    $ 38 "Switch JIG"
    switch_2 = JIG
    $ 39 "Case 1"
    if (1 == switch_2):
      $ 40 "3FG"
      $ 41 "define poses"
      $ 42 "FRM_Reference≔ULM_3FG"
      global FRM_Reference=ULM_3FG
      $ 43 "JNT_Q≔JNT_HOME"
      global JNT_Q=JNT_HOME
      $ 44 "PSE_T≔pose_trans(GRP_Offset, JIG_Offset)"
      global PSE_T= pose_trans (GRP_Offset, JIG_Offset)
      $ 45 "PSE_A≔pose_trans(PSE_T, p[0,0,0.100,0,0,0])"
      global PSE_A= pose_trans (PSE_T, p[0,0,0.100,0,0,0])
      $ 46 "PSE_R≔pose_add(PSE_T, p[0,0,0.100,0,0,0])"
      global PSE_R= pose_add (PSE_T, p[0,0,0.100,0,0,0])
    elif (2 == switch_2):
      $ 47 "Case 2"
      $ 48 "Input"
      $ 49 "'CHANGE THE REFERENCE TO THE FRAME TO MOVE IN'"
      # 'CHANGE THE REFERENCE TO THE FRAME TO MOVE IN'
      $ 50 "define poses"
      $ 51 "FRM_Reference≔ULM_Input"
      global FRM_Reference=ULM_Input
      $ 52 "PSE_T≔pose_trans(pose_trans(get_pattern_pos_rectangle(OBJ_Nbr, 'X', [10,5], patternsize=[0.181,0.081]), GRP_Offset), JIG_Offset)"
      global PSE_T= pose_trans ( pose_trans (get_pattern_pos_rectangle(OBJ_Nbr, "X", [10,5], patternsize=[0.181,0.081]), GRP_Offset), JIG_Offset)
      $ 53 "If Action≟1"
      if (Action == 1):
        $ 54 "PSE_R≔pose_add(PSE_T, p[0,0,0.200,0,0,0])"
        global PSE_R= pose_add (PSE_T, p[0,0,0.200,0,0,0])
        $ 55 "PSE_A≔pose_add(PSE_T, p[0,0,0.100,0,0,0])"
        global PSE_A= pose_add (PSE_T, p[0,0,0.100,0,0,0])
      else:
        $ 56 "ElseIf Action≟2"
        if (Action == 2):
          $ 57 "PSE_R≔pose_add(PSE_T, p[0,0,0.100,0,0,0])"
          global PSE_R= pose_add (PSE_T, p[0,0,0.100,0,0,0])
          $ 58 "PSE_A≔pose_add(PSE_T, p[0,0,0.200,0,0,0])"
          global PSE_A= pose_add (PSE_T, p[0,0,0.200,0,0,0])
        end
      end
    elif (3 == switch_2):
      $ 59 "Case 3"
      $ 60 "Output"
      $ 61 "'CHANGE THE REFERENCE TO THE FRAME TO MOVE IN'"
      # 'CHANGE THE REFERENCE TO THE FRAME TO MOVE IN'
      $ 62 "define poses"
      $ 63 "FRM_Reference≔ULM_Output"
      global FRM_Reference=ULM_Output
      $ 64 "PSE_T≔pose_trans(pose_trans(get_pattern_pos_rectangle(OBJ_Nbr, 'X', [10,5], patternsize=[0.181,0.081]), GRP_Offset), JIG_Offset)"
      global PSE_T= pose_trans ( pose_trans (get_pattern_pos_rectangle(OBJ_Nbr, "X", [10,5], patternsize=[0.181,0.081]), GRP_Offset), JIG_Offset)
      $ 66 "If Action≟1"
      if (Action == 1):
        $ 67 "PSE_R≔pose_add(PSE_T, p[0,0,0.200,0,0,0])"
        global PSE_R= pose_add (PSE_T, p[0,0,0.200,0,0,0])
        $ 68 "PSE_A≔pose_add(PSE_T, p[0,0,0.100,0,0,0])"
        global PSE_A= pose_add (PSE_T, p[0,0,0.100,0,0,0])
      else:
        $ 69 "ElseIf Action≟2"
        if (Action == 2):
          $ 70 "PSE_R≔pose_add(PSE_T, p[0,0,0.100,0,0,0])"
          global PSE_R= pose_add (PSE_T, p[0,0,0.100,0,0,0])
          $ 71 "PSE_A≔pose_add(PSE_T, p[0,0,0.200,0,0,0])"
          global PSE_A= pose_add (PSE_T, p[0,0,0.200,0,0,0])
        end
      end
    elif (4 == switch_2):
      $ 72 "Case 4"
      $ 73 "jig centrifuge racks"
      $ 74 "define poses"
      $ 75 "FRM_Reference≔ULM_Cent_Racks"
      global FRM_Reference=ULM_Cent_Racks
      $ 76 "PSE_T≔get_pattern_pos_rectangle(JIG_Slot, 'X', [4,1], patternsize=[0.291,0])"
      global PSE_T=get_pattern_pos_rectangle(JIG_Slot, "X", [4,1], patternsize=[0.291,0])
      $ 77 "If OBJ_Nbr≠0"
      if (OBJ_Nbr != 0):
        $ 78 "PSE_T≔pose_trans(pose_trans(PSE_T, get_pattern_pos_rectangle(OBJ_Nbr, 'X', [3,3], patternsize=[0.060,0.060])),p[-0.030, -0.030,0,0,0,3.927])"
        global PSE_T= pose_trans ( pose_trans (PSE_T, get_pattern_pos_rectangle(OBJ_Nbr, "X", [3,3], patternsize=[0.060,0.060])),p[-0.030, -0.030,0,0,0,3.927])
      end
      $ 79 "PSE_T≔pose_trans(PSE_T, GRP_Offset)"
      global PSE_T= pose_trans (PSE_T, GRP_Offset)
      $ 80 "If Action≟1"
      if (Action == 1):
        $ 81 "PSE_R≔pose_add(PSE_T, p[0,0,0.200,0,0,0])"
        global PSE_R= pose_add (PSE_T, p[0,0,0.200,0,0,0])
        $ 82 "PSE_A≔pose_add(PSE_T, p[0,0,0.100,0,0,0])"
        global PSE_A= pose_add (PSE_T, p[0,0,0.100,0,0,0])
      else:
        $ 83 "ElseIf Action≟2"
        if (Action == 2):
          $ 84 "PSE_R≔pose_add(PSE_T, p[0,0,0.100,0,0,0])"
          global PSE_R= pose_add (PSE_T, p[0,0,0.100,0,0,0])
          $ 85 "PSE_A≔pose_add(PSE_T, p[0,0,0.200,0,0,0])"
          global PSE_A= pose_add (PSE_T, p[0,0,0.200,0,0,0])
        end
      end
    end
  elif (2 == switch_1):
    $ 86 "Case 2"
    $ 87 "Centrifuge"
    $ 88 "'CHANGE THE REFERENCE TO THE FRAME TO MOVE IN'"
    # 'CHANGE THE REFERENCE TO THE FRAME TO MOVE IN'
    $ 89 "define poses"
    $ 90 "FRM_Reference≔FRM_Centrifuge"
    global FRM_Reference=FRM_Centrifuge
    $ 91 "PSE_T≔GRP_Offset"
    global PSE_T=GRP_Offset
    $ 92 "If Action≟8"
    if (Action == 8):
      $ 93 "PSE_R≔pose_add(PSE_T, p[0,0,0.250,0,0,0])"
      global PSE_R= pose_add (PSE_T, p[0,0,0.250,0,0,0])
      $ 94 "PSE_A≔pose_add(PSE_T, p[0,0,0.150,0,0,0])"
      global PSE_A= pose_add (PSE_T, p[0,0,0.150,0,0,0])
    else:
      $ 95 "ElseIf Action≟7"
      if (Action == 7):
        $ 96 "PSE_R≔pose_add(PSE_T, p[0,0,0.150,0,0,0])"
        global PSE_R= pose_add (PSE_T, p[0,0,0.150,0,0,0])
        $ 97 "PSE_A≔pose_add(PSE_T, p[0,0,0.250,0,0,0])"
        global PSE_A= pose_add (PSE_T, p[0,0,0.250,0,0,0])
      end
    end
  elif (3 == switch_1):
    $ 98 "Case 3"
    $ 99 "Output"
    $ 100 "'CHANGE THE REFERENCE TO THE FRAME TO MOVE IN'"
    # 'CHANGE THE REFERENCE TO THE FRAME TO MOVE IN'
    $ 101 "define poses"
    $ 102 "FRM_Reference≔Base_const"
    global FRM_Reference=p[0.0,0.0,0.0,0.0,0.0,0.0]
    $ 103 "PSE_T≔p[0,0,0,0,0,0]"
    global PSE_T=p[0,0,0,0,0,0]
    $ 104 "PSE_A≔pose_add(PSE_T, p[0,0,0.150,0,0,0])"
    global PSE_A= pose_add (PSE_T, p[0,0,0.150,0,0,0])
    $ 105 "PSE_R≔pose_add(PSE_T, p[0,0,0.100,0,0,0])"
    global PSE_R= pose_add (PSE_T, p[0,0,0.100,0,0,0])
  end
  $ 106 "Additional check"
  $ 107 "If  not is_reachable(FRM_Reference,[PSE_A,PSE_A_H,PSE_T,PSE_T_H,PSE_R,PSE_R_H])"
  if (  not  is_reachable(FRM_Reference,[PSE_A,PSE_A_H,PSE_T,PSE_T_H,PSE_R,PSE_R_H])):
    $ 108 "Error"
    $ 109 "set_error(ERROR_POSE_NOT_REACHABLE)"
    set_error(ERROR_POSE_NOT_REACHABLE)
    $ 110 "Action≔0"
    global Action=0
  end
  $ 111 "'=========='"
  # '=========='
  $ 112 "Switch Action"
  switch_1 = Action
  $ 113 "Case 1"
  if (1 == switch_1):
    $ 114 "Pick"
    $ 115 "Action_Info≔'pick object'"
    global Action_Info="pick object"
    $ 116 "do_transition(pose_trans(FRM_Reference, PSE_T), keep_rxry=OBJ_Picked)"
    do_transition( pose_trans (FRM_Reference, PSE_T), keep_rxry=OBJ_Picked)
    $ 117 "EOAT"
    $ 118 "If  not OBJ_Picked"
    if (  not  OBJ_Picked):
      $ 119 "rq_move_and_wait_mm(GRP_Open_Pos)"
       rq_move_and_wait_mm (GRP_Open_Pos)
    end
    $ 120 "If PSE_A_H≠PSE_Z"
    if (PSE_A_H != PSE_Z):
      $ 121 "If JNT_Q≠JNT_Z"
      if (JNT_Q != JNT_Z):
        $ 122 "movej(get_inverse_kin(pose_trans(FRM_Reference, PSE_A_H), qnear=JNT_Q), r=0.050)"
        movej(get_inverse_kin( pose_trans (FRM_Reference, PSE_A_H), qnear=JNT_Q), r=0.050)
      else:
        $ 123 "Else" "noBreak"
        $ 124 "movej(pose_trans(FRM_Reference, PSE_A_H), r=0.050)"
        movej( pose_trans (FRM_Reference, PSE_A_H), r=0.050)
      end
    end
    $ 125 "If PSE_A≠PSE_Z"
    if (PSE_A != PSE_Z):
      $ 126 "If JNT_Q≠JNT_Z"
      if (JNT_Q != JNT_Z):
        $ 127 "movej(get_inverse_kin(pose_trans(FRM_Reference, PSE_A), qnear=JNT_Q), r=0.020)"
        movej(get_inverse_kin( pose_trans (FRM_Reference, PSE_A), qnear=JNT_Q), r=0.020)
      else:
        $ 128 "Else" "noBreak"
        $ 129 "movej(pose_trans(FRM_Reference, PSE_A), r=0.020)"
        movej( pose_trans (FRM_Reference, PSE_A), r=0.020)
      end
    end
    $ 130 "MoveL"
    $ 131 "If PSE_T_H≠PSE_Z"
    if (PSE_T_H != PSE_Z):
      $ 132 "PSE_T_H" "breakAfter"
      movel(pose_trans(FRM_Reference, PSE_T_H), a=0.5, v=0.4, r=0.01)
    end
    $ 133 "PSE_T" "breakAfter"
    movel(pose_trans(FRM_Reference, PSE_T), a=0.08, v=0.12)
    $ 134 "EOAT"
    $ 135 "rq_set_force_norm(50)"
     rq_set_force_norm (50)
    $ 136 "rq_close_and_wait()"
     rq_close_and_wait ()
    $ 137 "OBJ_Picked≔rq_is_object_detected()"
    global OBJ_Picked= rq_is_object_detected ()
    $ 138 "If  not OBJ_Picked"
    if (  not  OBJ_Picked):
      $ 139 "set_error(ERROR_NO_OBJECT_TO_PICK)"
      set_error(ERROR_NO_OBJECT_TO_PICK)
    end
    $ 140 "EXTT"
    $ 141 "Switch JIG"
    switch_2 = JIG
    $ 142 "Case 1"
    if (1 == switch_2):
      $ 143 "3FG"
      $ 144 "If OBJ_Picked"
      if (OBJ_Picked):
        $ 145 "Set GRP_3F_Enable=On"
        set_standard_digital_out(4, True)
      end
    end
    $ 146 "If PSE_R_H≠PSE_Z"
    if (PSE_R_H != PSE_Z):
      $ 147 "PSE_R" "breakAfter"
      movel(pose_trans(FRM_Reference, PSE_R), a=0.5, v=0.4, r=0.01)
      $ 148 "PSE_R_H" "breakAfter"
      movel(pose_trans(FRM_Reference, PSE_R_H), a=0.5, v=0.4)
    else:
      $ 149 "Else" "noBreak"
      $ 150 "PSE_R" "breakAfter"
      movel(pose_trans(FRM_Reference, PSE_R), a=0.5, v=0.4)
    end
  elif (2 == switch_1):
    $ 151 "Case 2"
    $ 152 "Place"
    $ 153 "Action_Info≔'place object'"
    global Action_Info="place object"
    $ 154 "do_transition(pose_trans(FRM_Reference, PSE_T), keep_rxry=OBJ_Picked)"
    do_transition( pose_trans (FRM_Reference, PSE_T), keep_rxry=OBJ_Picked)
    $ 155 "EXTT"
    $ 156 "Switch JIG"
    switch_2 = JIG
    $ 157 "Case 1"
    if (1 == switch_2):
      $ 158 "3FG"
      $ 159 "If OBJ_Picked"
      if (OBJ_Picked):
        $ 160 "Set GRP_3F_Open=On"
        set_standard_digital_out(5, True)
      end
    end
    $ 161 "If PSE_A_H≠PSE_Z"
    if (PSE_A_H != PSE_Z):
      $ 162 "If JNT_Q≠JNT_Z"
      if (JNT_Q != JNT_Z):
        $ 163 "movej(get_inverse_kin(pose_trans(FRM_Reference, PSE_A_H), qnear=JNT_Q), r=0.050)"
        movej(get_inverse_kin( pose_trans (FRM_Reference, PSE_A_H), qnear=JNT_Q), r=0.050)
      else:
        $ 164 "Else" "noBreak"
        $ 165 "movej(pose_trans(FRM_Reference, PSE_A_H), r=0.050)"
        movej( pose_trans (FRM_Reference, PSE_A_H), r=0.050)
      end
    end
    $ 166 "If PSE_A≠PSE_Z"
    if (PSE_A != PSE_Z):
      $ 167 "If JNT_Q≠JNT_Z"
      if (JNT_Q != JNT_Z):
        $ 168 "movej(get_inverse_kin(pose_trans(FRM_Reference, PSE_A), qnear=JNT_Q), r=0.020)"
        movej(get_inverse_kin( pose_trans (FRM_Reference, PSE_A), qnear=JNT_Q), r=0.020)
      else:
        $ 169 "Else" "noBreak"
        $ 170 "movej(pose_trans(FRM_Reference, PSE_A), r=0.020)"
        movej( pose_trans (FRM_Reference, PSE_A), r=0.020)
      end
    end
    $ 171 "MoveL"
    $ 172 "If PSE_T_H≠PSE_Z"
    if (PSE_T_H != PSE_Z):
      $ 173 "PSE_T_H" "breakAfter"
      movel(pose_trans(FRM_Reference, PSE_T_H), a=0.5, v=0.4, r=0.01)
    end
    $ 174 "PSE_T" "breakAfter"
    global move_thread_flag_174=0
    thread move_thread_174():
      enter_critical
      move_thread_flag_174 = 1
      movel(pose_trans(FRM_Reference, PSE_T), a=0.05, v=0.09)
      move_thread_flag_174 = 2
      exit_critical
    end
    move_thread_flag_174 = 0
    move_thread_han_174 = run move_thread_174()
    while (True):
      local targetTcpDirection=get_target_tcp_speed()
      local stepsToRetract=tool_contact(direction=targetTcpDirection)
      if (stepsToRetract > 0):
        kill move_thread_han_174
        stopl(0.5)
        $ 175 "Until (tool_contact_detection)"
        break
      end
      sleep(1.0E-10)
      if (move_thread_flag_174 > 1):
        join move_thread_han_174
        break
      end
      sync()
    end
    $ 176 "Force"
    sleep(0.02)
    zero_ftsensor()
    force_mode(FRM_Reference, [1, 1, 1, 0, 0, 0], [0.0, 0.0, 0.0, 0.0, 0.0, 0.0], 2, [0.1, 0.1, 0.01, 0.3490658503988659, 0.3490658503988659, 0.3490658503988659])
    $ 177 "PSE_T" "noBreak"
    movel(pose_trans(FRM_Reference, PSE_T), a=0.04, v=0.07)
    end_force_mode()
    stopl(5.0)
    $ 178 "EXTT"
    $ 179 "Switch JIG"
    switch_2 = JIG
    $ 180 "Case 1"
    if (1 == switch_2):
      $ 181 "3FG"
      $ 182 "If OBJ_Picked"
      if (OBJ_Picked):
        $ 183 "Set GRP_3F_Open=Off"
        set_standard_digital_out(5, False)
        $ 184 "Wait: 0.2"
        sleep(0.2)
      end
    end
    $ 185 "EOAT"
    $ 186 "rq_move_and_wait_mm(GRP_Open_Pos)"
     rq_move_and_wait_mm (GRP_Open_Pos)
    $ 187 "OBJ_Picked≔rq_is_object_detected()"
    global OBJ_Picked= rq_is_object_detected ()
    $ 188 "If PSE_R_H≠PSE_Z"
    if (PSE_R_H != PSE_Z):
      $ 189 "PSE_R" "breakAfter"
      movel(pose_trans(FRM_Reference, PSE_R), a=0.5, v=0.4, r=0.01)
      $ 190 "PSE_R_H" "breakAfter"
      movel(pose_trans(FRM_Reference, PSE_R_H), a=0.5, v=0.4)
    else:
      $ 191 "Else" "noBreak"
      $ 192 "PSE_R" "breakAfter"
      movel(pose_trans(FRM_Reference, PSE_R), a=0.5, v=0.4)
    end
  elif (3 == switch_1):
    $ 193 "Case 3"
    $ 194 "Push"
    $ 195 "Action_Info≔'push'"
    global Action_Info="push"
  elif (4 == switch_1):
    $ 196 "Case 4"
    $ 197 "Pull"
    $ 198 "Action_Info≔'pull'"
    global Action_Info="pull"
  elif (7 == switch_1):
    $ 199 "Case 7"
    $ 200 "Load"
    $ 201 "Action_Info≔'load object'"
    global Action_Info="load object"
    $ 202 "do_transition(pose_trans(FRM_Reference, PSE_T), keep_rxry=OBJ_Picked)"
    do_transition( pose_trans (FRM_Reference, PSE_T), keep_rxry=OBJ_Picked)
    $ 203 "If PSE_A_H≠PSE_Z"
    if (PSE_A_H != PSE_Z):
      $ 204 "If JNT_Q≠JNT_Z"
      if (JNT_Q != JNT_Z):
        $ 205 "movej(get_inverse_kin(pose_trans(FRM_Reference, PSE_A_H), qnear=JNT_Q), r=0.050)"
        movej(get_inverse_kin( pose_trans (FRM_Reference, PSE_A_H), qnear=JNT_Q), r=0.050)
      else:
        $ 206 "Else" "noBreak"
        $ 207 "movej(pose_trans(FRM_Reference, PSE_A_H), r=0.050)"
        movej( pose_trans (FRM_Reference, PSE_A_H), r=0.050)
      end
    end
    $ 208 "If PSE_A≠PSE_Z"
    if (PSE_A != PSE_Z):
      $ 209 "If JNT_Q≠JNT_Z"
      if (JNT_Q != JNT_Z):
        $ 210 "movej(get_inverse_kin(pose_trans(FRM_Reference, PSE_A), qnear=JNT_Q), r=0.020)"
        movej(get_inverse_kin( pose_trans (FRM_Reference, PSE_A), qnear=JNT_Q), r=0.020)
      else:
        $ 211 "Else" "noBreak"
        $ 212 "movej(pose_trans(FRM_Reference, PSE_A), r=0.020)"
        movej( pose_trans (FRM_Reference, PSE_A), r=0.020)
      end
    end
    $ 213 "MoveL"
    $ 214 "If PSE_T_H≠PSE_Z"
    if (PSE_T_H != PSE_Z):
      $ 215 "PSE_T_H" "breakAfter"
      movel(pose_trans(FRM_Reference, PSE_T_H), a=0.5, v=0.4, r=0.01)
    end
    $ 216 "PSE_T" "breakAfter"
    global move_thread_flag_216=0
    thread move_thread_216():
      enter_critical
      move_thread_flag_216 = 1
      movel(pose_trans(FRM_Reference, PSE_T), a=0.05, v=0.09)
      move_thread_flag_216 = 2
      exit_critical
    end
    move_thread_flag_216 = 0
    move_thread_han_216 = run move_thread_216()
    while (True):
      local targetTcpDirection=get_target_tcp_speed()
      local stepsToRetract=tool_contact(direction=targetTcpDirection)
      if (stepsToRetract > 0):
        kill move_thread_han_216
        stopl(0.5)
        $ 217 "Until (tool_contact_detection)"
        break
      end
      sleep(1.0E-10)
      if (move_thread_flag_216 > 1):
        join move_thread_han_216
        break
      end
      sync()
    end
    $ 218 "Force"
    sleep(0.02)
    zero_ftsensor()
    force_mode(FRM_Reference, [0, 1, 1, 0, 0, 1], [0.0, 0.0, 0.0, 0.0, 0.0, 0.0], 2, [0.1, 0.05, 0.02, 0.3490658503988659, 0.3490658503988659, 3.141592653589793])
    $ 219 "PSE_T" "noBreak"
    movel(pose_trans(FRM_Reference, PSE_T), a=0.04, v=0.07)
    end_force_mode()
    stopl(5.0)
    $ 220 "EOAT"
    $ 221 "rq_move_and_wait_mm(GRP_Open_Pos)"
     rq_move_and_wait_mm (GRP_Open_Pos)
    $ 222 "OBJ_Picked≔rq_is_object_detected()"
    global OBJ_Picked= rq_is_object_detected ()
    $ 223 "If PSE_R_H≠PSE_Z"
    if (PSE_R_H != PSE_Z):
      $ 224 "PSE_R" "breakAfter"
      movel(pose_trans(FRM_Reference, PSE_R), a=0.5, v=0.4, r=0.01)
      $ 225 "PSE_R_H" "breakAfter"
      movel(pose_trans(FRM_Reference, PSE_R_H), a=0.5, v=0.4)
    else:
      $ 226 "Else" "noBreak"
      $ 227 "PSE_R" "breakAfter"
      movel(pose_trans(FRM_Reference, PSE_R), a=0.5, v=0.4)
    end
  elif (8 == switch_1):
    $ 228 "Case 8"
    $ 229 "Unload"
    $ 230 "Action_Info≔'pick object'"
    global Action_Info="pick object"
    $ 231 "do_transition(pose_trans(FRM_Reference, PSE_T), keep_rxry=OBJ_Picked)"
    do_transition( pose_trans (FRM_Reference, PSE_T), keep_rxry=OBJ_Picked)
    $ 232 "EOAT"
    $ 233 "If  not OBJ_Picked"
    if (  not  OBJ_Picked):
      $ 234 "rq_move_and_wait_mm(GRP_Open_Pos)"
       rq_move_and_wait_mm (GRP_Open_Pos)
    end
    $ 235 "If PSE_A_H≠PSE_Z"
    if (PSE_A_H != PSE_Z):
      $ 236 "If JNT_Q≠JNT_Z"
      if (JNT_Q != JNT_Z):
        $ 237 "movej(get_inverse_kin(pose_trans(FRM_Reference, PSE_A_H), qnear=JNT_Q), r=0.050)"
        movej(get_inverse_kin( pose_trans (FRM_Reference, PSE_A_H), qnear=JNT_Q), r=0.050)
      else:
        $ 238 "Else" "noBreak"
        $ 239 "movej(pose_trans(FRM_Reference, PSE_A_H), r=0.050)"
        movej( pose_trans (FRM_Reference, PSE_A_H), r=0.050)
      end
    end
    $ 240 "If PSE_A≠PSE_Z"
    if (PSE_A != PSE_Z):
      $ 241 "If JNT_Q≠JNT_Z"
      if (JNT_Q != JNT_Z):
        $ 242 "movej(get_inverse_kin(pose_trans(FRM_Reference, PSE_A), qnear=JNT_Q), r=0.020)"
        movej(get_inverse_kin( pose_trans (FRM_Reference, PSE_A), qnear=JNT_Q), r=0.020)
      else:
        $ 243 "Else" "noBreak"
        $ 244 "movej(pose_trans(FRM_Reference, PSE_A), r=0.020)"
        movej( pose_trans (FRM_Reference, PSE_A), r=0.020)
      end
    end
    $ 245 "MoveL"
    $ 246 "If PSE_T_H≠PSE_Z"
    if (PSE_T_H != PSE_Z):
      $ 247 "PSE_T_H" "breakAfter"
      movel(pose_trans(FRM_Reference, PSE_T_H), a=0.5, v=0.4, r=0.01)
    end
    $ 248 "PSE_T" "breakAfter"
    movel(pose_trans(FRM_Reference, PSE_T), a=0.08, v=0.12)
    $ 249 "Force"
    sleep(0.02)
    zero_ftsensor()
    force_mode(FRM_Reference, [1, 1, 0, 0, 0, 0], [0.0, 0.0, 0.0, 0.0, 0.0, 0.0], 2, [0.05, 0.05, 0.1, 0.3490658503988659, 0.3490658503988659, 0.3490658503988659])
    $ 250 "EOAT" "noBreak"
    $ 251 "rq_set_force_norm(50)" "noBreak"
     rq_set_force_norm (50)
    $ 252 "rq_close_and_wait()" "noBreak"
     rq_close_and_wait ()
    $ 253 "OBJ_Picked≔rq_is_object_detected()" "noBreak"
    global OBJ_Picked= rq_is_object_detected ()
    $ 254 "If  not OBJ_Picked" "noBreak"
    if (  not  OBJ_Picked):
      $ 255 "set_error(ERROR_NO_OBJECT_TO_PICK)" "noBreak"
      set_error(ERROR_NO_OBJECT_TO_PICK)
    end
    $ 256 "If PSE_R_H≠PSE_Z" "noBreak"
    if (PSE_R_H != PSE_Z):
      $ 257 "PSE_R" "noBreak"
      movel(pose_trans(FRM_Reference, PSE_R), a=0.5, v=0.4, r=0.01)
      $ 258 "PSE_R_H" "noBreak"
      movel(pose_trans(FRM_Reference, PSE_R_H), a=0.5, v=0.4)
    else:
      $ 259 "Else" "noBreak"
      $ 260 "PSE_R" "noBreak"
      movel(pose_trans(FRM_Reference, PSE_R), a=0.5, v=0.4)
    end
    end_force_mode()
    stopl(5.0)
  elif (12 == switch_1):
    $ 261 "Case 12"
    $ 262 "Decap"
    $ 263 "Action_Info≔'decapping'"
    global Action_Info="decapping"
    $ 264 "Set GRP_3F_Enable=On"
    set_standard_digital_out(4, True)
    $ 265 "Set GRP_3F_Decap=On"
    set_standard_digital_out(3, True)
    $ 266 "Force"
    sleep(0.02)
    zero_ftsensor()
    force_mode(tool_pose(), [0, 0, 1, 0, 0, 0], [0.0, 0.0, 5.0, 0.0, 0.0, 0.0], 2, [0.1, 0.1, 0.15, 0.3490658503988659, 0.3490658503988659, 0.3490658503988659])
    $ 267 "check_decapping(offset=0.015, timeout=5, abort=CMD_Hold)" "noBreak"
    check_decapping(offset=0.015, timeout=5, abort=CMD_Hold)
    end_force_mode()
    stopl(5.0)
    $ 268 "Set GRP_3F_Decap=Off"
    set_standard_digital_out(3, False)
    $ 269 "Set GRP_3F_Enable=Off"
    set_standard_digital_out(4, False)
    $ 270 "MoveL"
    $ 271 "PSE_R" "breakAfter"
    movel(pose_trans(FRM_Reference, PSE_R), a=0.8, v=0.15)
  elif (13 == switch_1):
    $ 272 "Case 13"
    $ 273 "Read"
    $ 274 "Preorient"
    $ 275 "TMR_Barcode: Reset"
    TMR_Barcode = 0
    $ 276 "Set BarcodeTrigger=HI:Pulse 0.1"
    thread SinglePulse2():
      set_standard_digital_out(6, True)
      sleep(0.1)
      set_standard_digital_out(6, False)
    end
    singlePulse2 = run SinglePulse2()
    $ 277 "Wait Barcode_OK or Barcode_nOK"
    while (not(get_standard_digital_in(6)  or  get_standard_digital_in(7))):
      sync()
    end
    $ 278 "If Barcode_OK"
    if (get_standard_digital_in(6)):
      $ 279 "Set GRP_3F_Decap=HI:Pulse 2.0"
      thread SinglePulse3():
        set_standard_digital_out(3, True)
        sleep(2.0)
        set_standard_digital_out(3, False)
      end
      singlePulse3 = run SinglePulse3()
    end
    $ 280 "Search for code"
    $ 281 "Wait ( not Barcode_OK and  not Barcode_nOK and  not GRP_3F_Decap)"
    while (not((  not  get_standard_digital_in(6)  and    not  get_standard_digital_in(7)  and    not  get_standard_digital_out(3)))):
      sync()
    end
    $ 282 "TMR_Barcode: Start"
    TMR_Barcode_is_counting = True
    $ 283 "Set GRP_3F_Cap=On"
    set_standard_digital_out(2, True)
    $ 284 "Set BarcodeTrigger=On"
    set_standard_digital_out(6, True)
    $ 285 "Wait TMR_Barcode≥PRM_TO_Read_BC or Barcode_OK or Barcode_nOK"
    while (not(TMR_Barcode >= PRM_TO_Read_BC  or  get_standard_digital_in(6)  or  get_standard_digital_in(7))):
      sync()
    end
    $ 286 "Set GRP_3F_Cap=Off"
    set_standard_digital_out(2, False)
    $ 287 "Set BarcodeTrigger=Off"
    set_standard_digital_out(6, False)
    $ 288 "TMR_Barcode: Stop"
    TMR_Barcode_is_counting = False
    $ 289 "If Barcode_OK"
    if (get_standard_digital_in(6)):
      $ 290 "barcode found"
      $ 291 "'nothing'"
      # 'nothing'
    else:
      $ 292 "ElseIf Barcode_nOK or TMR_Barcode≥PRM_TO_Read_BC"
      if (get_standard_digital_in(7)  or  TMR_Barcode >= PRM_TO_Read_BC):
        $ 293 "exeption"
        $ 294 "error"
        $ 295 "set_error(6000)"
        set_error(6000)
      end
    end
  elif (15 == switch_1):
    $ 296 "Case 15"
    $ 297 "Detect"
    $ 298 "Action_Info≔'detect'"
    global Action_Info="detect"
  end
  $ 299 "'=========='"
  # '=========='
  $ 300 "PostSettings"
  $ 301 "'ADD ADDITIONAL CHECKS'"
  # 'ADD ADDITIONAL CHECKS'
end
